Fanuc KAREL source: KO00061.KL

PROGRAM KO00061
%NOLOCKGROUP
%ENVIRONMENT MIR
VAR
  P1: XYZWPR
  P2: JOINTPOS
  F: BOOLEAN
  OUT: POSITION
BEGIN
  F = TRUE
  OUT = MIRROR(P1, P2, F)
END KO00061
